FUNCTION_BLOCK RecoveryComposite (* Recoverable importer normalization cases *)
  (* Standard: 61499-1; Description: Copyright (c) 2026 Martin Erich Jobst This program and the accompanying materials are made available under the terms of the Eclipse Public License 2.0 which is available at https://www.eclipse.org/legal/epl-2.0/ SPDX-License-Identifier: EPL-2.0 *)
  (* Version 1.0, 2026-10-23, Martin Jobst *)
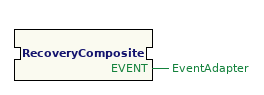
  PLUGS
    EVENT : EventAdapter; (* Event/data adapter *) {SET_ATTRIBUTE(AdapterAttribute, AdapterValue)} {SET_ATTRIBUTE(PinComment, REQD:legacy adapter pin comment)} {SET_ATTRIBUTE(VarConfig, REQD:true)}
  END_PLUGS
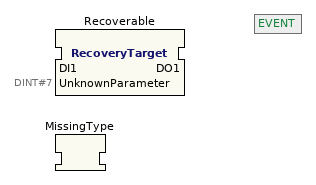
  FBS
    Recoverable : RecoveryTarget(UnknownParameter := DINT#7); {SET_ATTRIBUTE(Retain, TRUE)} {SET_ATTRIBUTE(PinComment, DI1:legacy input comment)} {SET_ATTRIBUTE(VarConfig, DI1:true)}
    MissingType : ;
  END_FBS
END_FUNCTION_BLOCK
